// TIA Portal V21 export
FUNCTION_BLOCK "F_FB_MainSafety"   // FB3, F_LAD
{ S7_Optimized_Access := 'TRUE' }
   VAR
      Enable : Bool;   // Schutztür geschlossen und Not-Halt in Ordnung / Guard closed and emergency stop ok
      Released : Bool;   // Maschine freigegeben / Machine released
      LogicRelease : Bool;   // Freigabe aus F_FC_Logic / Release from F_FC_Logic
   END_VAR
BEGIN

REGION Network 1: F-DB lesen / Read the F-DB
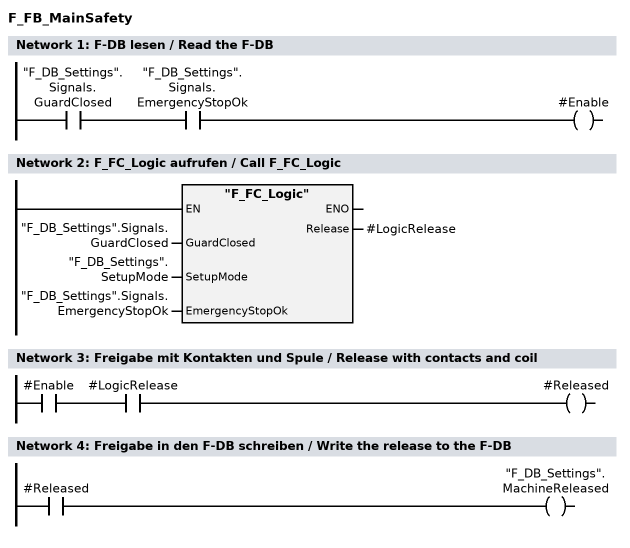
   RUNG wire#powerrail
      Contact( "F_DB_Settings".Signals.GuardClosed )
      Contact( "F_DB_Settings".Signals.EmergencyStopOk )
      Coil( #Enable )
   END_RUNG
   // the same network as SCL:
   #Enable := "F_DB_Settings".Signals.GuardClosed AND "F_DB_Settings".Signals.EmergencyStopOk;
END_REGION

REGION Network 2: F_FC_Logic aufrufen / Call F_FC_Logic
   RUNG wire#powerrail
      "F_FC_Logic"(GuardClosed := "F_DB_Settings".Signals.GuardClosed, SetupMode := "F_DB_Settings".SetupMode, EmergencyStopOk := "F_DB_Settings".Signals.EmergencyStopOk, Release => #LogicRelease)
   END_RUNG
   // the same network as SCL:
   "F_FC_Logic"(GuardClosed := "F_DB_Settings".Signals.GuardClosed,
                SetupMode := "F_DB_Settings".SetupMode,
                EmergencyStopOk := "F_DB_Settings".Signals.EmergencyStopOk,
                Release => #LogicRelease);
END_REGION

REGION Network 3: Freigabe mit Kontakten und Spule / Release with contacts and coil
   RUNG wire#powerrail
      Contact( #Enable )
      Contact( #LogicRelease )
      Coil( #Released )
   END_RUNG
   // the same network as SCL:
   #Released := #Enable AND #LogicRelease;
END_REGION

REGION Network 4: Freigabe in den F-DB schreiben / Write the release to the F-DB
   RUNG wire#powerrail
      Contact( #Released )
      Coil( "F_DB_Settings".MachineReleased )
   END_RUNG
   // the same network as SCL:
   "F_DB_Settings".MachineReleased := #Released;
END_REGION
END_FUNCTION_BLOCK
